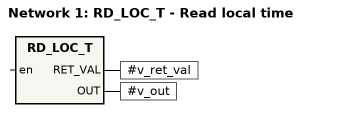
   #v_ret_val := RD_LOC_T(OUT => #v_out);
END_REGION
END_FUNCTION_BLOCK

FUNCTION_BLOCK "FB_Fbd_ex011"   // FB73, FBD
{ S7_Optimized_Access := 'TRUE' }
   VAR_INPUT
      v_req : Bool;
      v_timezone : TimeTransformationRule;
   END_VAR
   VAR_OUTPUT
      v_done : Bool;
      v_busy : Bool;
      v_error : Bool;
      v_status : Word;
   END_VAR
   VAR
      inst : SET_TIMEZONE;
   END_VAR
BEGIN

REGION Network 1: SET_TIMEZONE - Set time zone
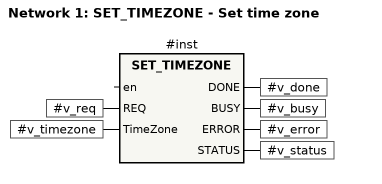
   #inst(REQ := #v_req,   // SET_TIMEZONE
         TimeZone := #v_timezone,
         DONE => #v_done,
         BUSY => #v_busy,
         ERROR => #v_error,
         STATUS => #v_status);
END_REGION
END_FUNCTION_BLOCK

FUNCTION_BLOCK "FB_Fbd_ex012"   // FB74, FBD
{ S7_Optimized_Access := 'TRUE' }
   VAR_OUTPUT
      v_ret_val : Int;
   END_VAR
BEGIN

REGION Network 1: SNC_RTCB - Synchronize slave clocks
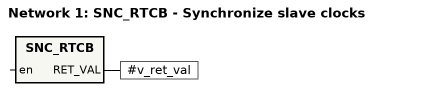
   #v_ret_val := SNC_RTCB();
END_REGION
END_FUNCTION_BLOCK

FUNCTION_BLOCK "FB_Fbd_ex013"   // FB75, FBD
{ S7_Optimized_Access := 'TRUE' }
   VAR_OUTPUT
      v_ret_val : Time;
   END_VAR
BEGIN

REGION Network 1: TIME_TCK - Read time counter
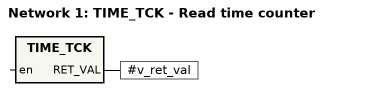
   #v_ret_val := TIME_TCK();
END_REGION
END_FUNCTION_BLOCK

FUNCTION_BLOCK "FB_Fbd_ex014"   // FB76, FBD
{ S7_Optimized_Access := 'TRUE' }
   VAR_INPUT
      v_nr : Rtm;
      v_mode : Byte;
      v_pv : DInt;
   END_VAR
   VAR_OUTPUT
      v_ret_val : Int;
      v_cq : Bool;
      v_cv : DInt;
   END_VAR
BEGIN

REGION Network 1: RTM - Runtime meters
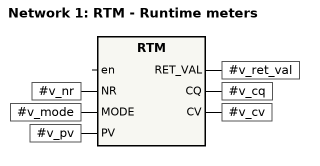
   #v_ret_val := RTM(NR := #v_nr, MODE := #v_mode, PV := #v_pv, CQ => #v_cq, CV => #v_cv);
END_REGION
END_FUNCTION_BLOCK

FUNCTION_BLOCK "FB_Fbd_ex015"   // FB77, FBD
{ S7_Optimized_Access := 'TRUE' }
   VAR_INPUT
      v_in : String;
   END_VAR
   VAR_OUTPUT
      v_out : String;
   END_VAR
BEGIN

REGION Network 1: S_MOVE - Move character string
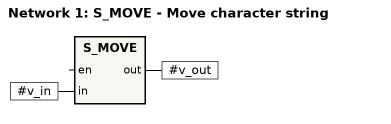
   #v_out := #v_in;
END_REGION
END_FUNCTION_BLOCK

FUNCTION_BLOCK "FB_Fbd_ex025"   // FB78, FBD
{ S7_Optimized_Access := 'TRUE' }
   VAR_INPUT
      v_n : Int;
   END_VAR
   VAR_OUTPUT
      v_ret_val : Word;
   END_VAR
   VAR_IN_OUT
      v_in : Variant;
      v_out : Variant;
   END_VAR
BEGIN

REGION Network 1: ATH - Convert ASCII string to hexadecimal number
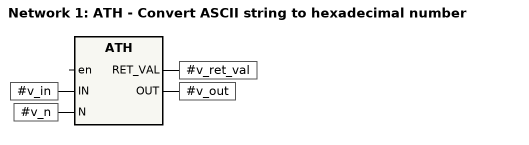
   #v_ret_val := ATH(IN := #v_in, N := #v_n, OUT => #v_out);
END_REGION
END_FUNCTION_BLOCK

FUNCTION_BLOCK "FB_Fbd_ex026"   // FB79, FBD
{ S7_Optimized_Access := 'TRUE' }
   VAR_INPUT
      v_n : UInt;
   END_VAR
   VAR_OUTPUT
      v_ret_val : Word;
   END_VAR
   VAR_IN_OUT
      v_in : Variant;
      v_out : Variant;
   END_VAR
BEGIN

REGION Network 1: HTA - Convert hexadecimal number to ASCII string
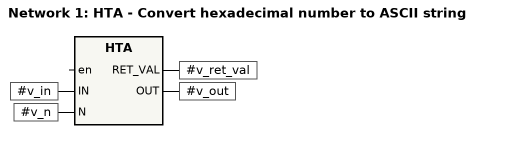
   #v_ret_val := HTA(IN := #v_in, N := #v_n, OUT => #v_out);
END_REGION
END_FUNCTION_BLOCK

FUNCTION_BLOCK "FB_Fbd_ex036"   // FB80, FBD
{ S7_Optimized_Access := 'TRUE' }
   VAR_INPUT
      v_size : DInt;
   END_VAR
   VAR_OUTPUT
      v_out : WString;
   END_VAR
   VAR_IN_OUT
      v_variable : Variant;
   END_VAR
BEGIN

REGION Network 1: GetSymbolName - Read out a tag on the input parameter
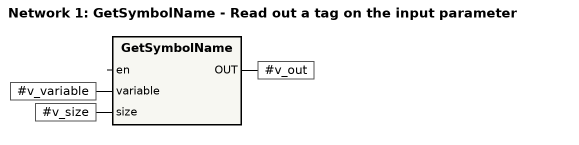
   // no SCL statement known for GetSymbolName: written as a call
   #v_out := GetSymbolName(variable := #v_variable, size := #v_size);
END_REGION
END_FUNCTION_BLOCK

FUNCTION_BLOCK "FB_Fbd_ex038"   // FB81, FBD
{ S7_Optimized_Access := 'TRUE' }
   VAR_INPUT
      v_size : DInt;
   END_VAR
   VAR_OUTPUT
      v_out : WString;
   END_VAR
BEGIN

REGION Network 1: GetInstanceName - Read out name of the read instance
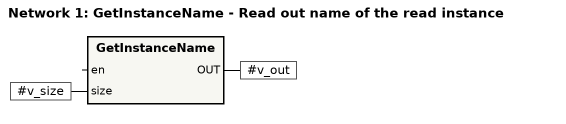
   // no SCL statement known for GetInstanceName: written as a call
   #v_out := GetInstanceName(size := #v_size);
END_REGION
END_FUNCTION_BLOCK

FUNCTION_BLOCK "FB_Fbd_ex039"   // FB82, FBD
{ S7_Optimized_Access := 'TRUE' }
   VAR_INPUT
      v_size : DInt;
   END_VAR
   VAR_OUTPUT
      v_out : WString;
   END_VAR
BEGIN

REGION Network 1: GetInstancePath - Query composite global name of the block instance
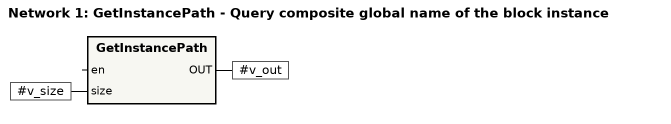
   // no SCL statement known for GetInstancePath: written as a call
   #v_out := GetInstancePath(size := #v_size);
END_REGION
END_FUNCTION_BLOCK

FUNCTION_BLOCK "FB_Fbd_ex040"   // FB83, FBD
{ S7_Optimized_Access := 'TRUE' }
   VAR_INPUT
      v_size : DInt;
   END_VAR
   VAR_OUTPUT
      v_ret_val : WString;
   END_VAR
BEGIN

REGION Network 1: GetBlockName - Read out name of the block
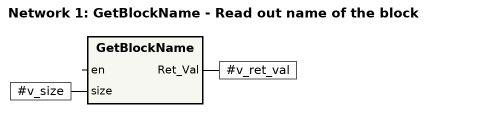
   // no SCL statement known for GetBlockName: written as a call
   #v_ret_val := GetBlockName(size := #v_size);
END_REGION
END_FUNCTION_BLOCK

FUNCTION_BLOCK "FB_Fbd_ex041"   // FB84, FBD
{ S7_Optimized_Access := 'TRUE' }
   VAR_INPUT
      v_part : Pip;
   END_VAR
   VAR_OUTPUT
      v_ret_val : Int;
      v_fladdr : Word;
   END_VAR
BEGIN

REGION Network 1: UPDAT_PI - Update the process image inputs
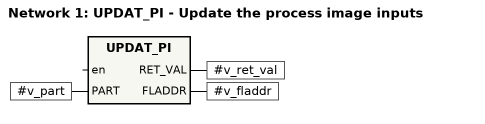
   #v_ret_val := UPDAT_PI(PART := #v_part, FLADDR => #v_fladdr);
END_REGION
END_FUNCTION_BLOCK

FUNCTION_BLOCK "FB_Fbd_ex042"   // FB85, FBD
{ S7_Optimized_Access := 'TRUE' }
   VAR_INPUT
      v_part : Pip;
   END_VAR
   VAR_OUTPUT
      v_ret_val : Int;
      v_fladdr : Word;
   END_VAR
BEGIN

REGION Network 1: UPDAT_PO - Update the process image outputs
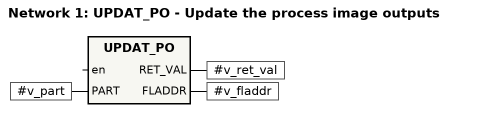
   #v_ret_val := UPDAT_PO(PART := #v_part, FLADDR => #v_fladdr);
END_REGION
END_FUNCTION_BLOCK

FUNCTION_BLOCK "FB_Fbd_ex043"   // FB86, FBD
{ S7_Optimized_Access := 'TRUE' }
   VAR_INPUT
      v_part : Pip;
   END_VAR
   VAR_OUTPUT
      v_ret_val : Int;
      v_fladdr : Word;
   END_VAR
BEGIN

REGION Network 1: SYNC_PI - Synchronize the process image inputs
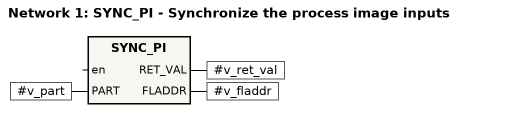
   #v_ret_val := SYNC_PI(PART := #v_part, FLADDR => #v_fladdr);
END_REGION
END_FUNCTION_BLOCK

FUNCTION_BLOCK "FB_Fbd_ex044"   // FB87, FBD
{ S7_Optimized_Access := 'TRUE' }
   VAR_INPUT
      v_part : Pip;
   END_VAR
   VAR_OUTPUT
      v_ret_val : Int;
      v_fladdr : Word;
   END_VAR
BEGIN

REGION Network 1: SYNC_PO - Synchronize the process image outputs
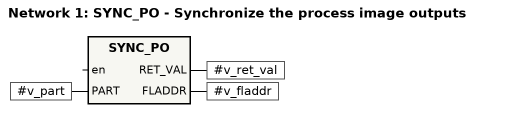
   #v_ret_val := SYNC_PO(PART := #v_part, FLADDR => #v_fladdr);
END_REGION
END_FUNCTION_BLOCK

FUNCTION_BLOCK "FB_Fbd_ex045"   // FB88, FBD
{ S7_Optimized_Access := 'TRUE' }
   VAR_INPUT
      v_req : Bool;
      v_id : Hw_Io;
      v_index : DInt;
      v_mlen : UInt;
   END_VAR
   VAR_OUTPUT
      v_valid : Bool;
      v_busy : Bool;
      v_error : Bool;
      v_status : DWord;
      v_len : UInt;
   END_VAR
   VAR_IN_OUT
      v_record : Array[0..99] of Byte;
   END_VAR
   VAR
      inst : RDREC;
   END_VAR
BEGIN

REGION Network 1: RDREC - Read data record
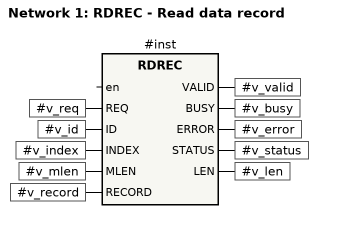
   #inst(REQ := #v_req,   // RDREC
         ID := #v_id,
         INDEX := #v_index,
         MLEN := #v_mlen,
         RECORD := #v_record,
         VALID => #v_valid,
         BUSY => #v_busy,
         ERROR => #v_error,
         STATUS => #v_status,
         LEN => #v_len);
END_REGION
END_FUNCTION_BLOCK

FUNCTION_BLOCK "FB_Fbd_ex046"   // FB89, FBD
{ S7_Optimized_Access := 'TRUE' }
   VAR_INPUT
      v_req : Bool;
      v_id : Hw_Io;
      v_index : DInt;
      v_len : UInt;
   END_VAR
   VAR_OUTPUT
      v_done : Bool;
      v_busy : Bool;
      v_error : Bool;
      v_status : DWord;
   END_VAR
   VAR_IN_OUT
      v_record : Array[0..99] of Byte;
   END_VAR
   VAR
      inst : WRREC;
   END_VAR
BEGIN

REGION Network 1: WRREC - Write data record
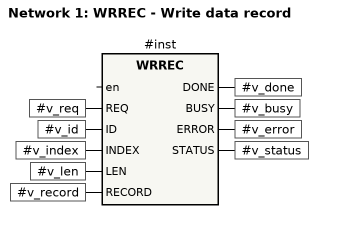
   #inst(REQ := #v_req,   // WRREC
         ID := #v_id,
         INDEX := #v_index,
         LEN := #v_len,
         RECORD := #v_record,
         DONE => #v_done,
         BUSY => #v_busy,
         ERROR => #v_error,
         STATUS => #v_status);
END_REGION
END_FUNCTION_BLOCK

FUNCTION_BLOCK "FB_Fbd_ex047"   // FB90, FBD
{ S7_Optimized_Access := 'TRUE' }
   VAR_INPUT
      v_id : Hw_SubModule;
   END_VAR
   VAR_OUTPUT
      v_status : DWord;
      v_len : Int;
   END_VAR
   VAR_IN_OUT
      v_inputs : Array[0..99] of Byte;
   END_VAR
   VAR
      inst : GETIO;
   END_VAR
BEGIN

REGION Network 1: GETIO - Read all inputs of a submodule
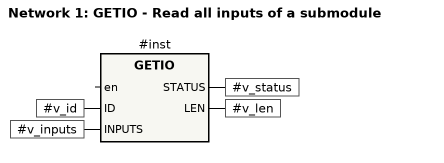
   #inst(ID := #v_id, INPUTS := #v_inputs, STATUS => #v_status, LEN => #v_len);   // GETIO
END_REGION
END_FUNCTION_BLOCK

FUNCTION_BLOCK "FB_Fbd_ex048"   // FB91, FBD
{ S7_Optimized_Access := 'TRUE' }
   VAR_INPUT
      v_id : Hw_SubModule;
   END_VAR
   VAR_OUTPUT
      v_status : DWord;
   END_VAR
   VAR_IN_OUT
      v_outputs : Array[0..99] of Byte;
   END_VAR
   VAR
      inst : SETIO;
   END_VAR
BEGIN

REGION Network 1: SETIO - Write all outputs of a submodule
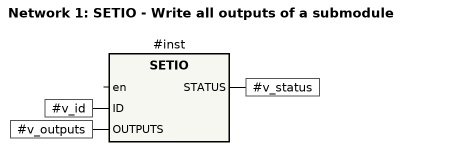
   #inst(ID := #v_id, OUTPUTS := #v_outputs, STATUS => #v_status);   // SETIO
END_REGION
END_FUNCTION_BLOCK

FUNCTION_BLOCK "FB_Fbd_ex049"   // FB92, FBD
{ S7_Optimized_Access := 'TRUE' }
   VAR_INPUT
      v_id : Hw_SubModule;
      v_offset : Int;
      v_len : Int;
   END_VAR
   VAR_OUTPUT
      v_status : DWord;
      v_error : Bool;
   END_VAR
   VAR_IN_OUT
      v_inputs : Array[0..99] of Byte;
   END_VAR
   VAR
      inst : GETIO_PART;
   END_VAR
BEGIN

REGION Network 1: GETIO_PART - Read inputs of a submodule
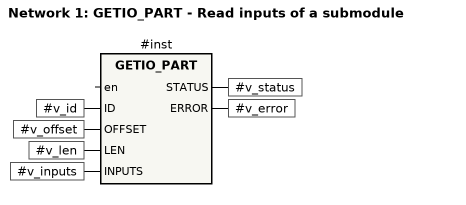
   #inst(ID := #v_id,   // GETIO_PART
         OFFSET := #v_offset,
         LEN := #v_len,
         INPUTS := #v_inputs,
         STATUS => #v_status,
         ERROR => #v_error);
END_REGION
END_FUNCTION_BLOCK

FUNCTION_BLOCK "FB_Fbd_ex050"   // FB93, FBD
{ S7_Optimized_Access := 'TRUE' }
   VAR_INPUT
      v_id : Hw_SubModule;
      v_offset : Int;
      v_len : Int;
   END_VAR
   VAR_OUTPUT
      v_status : DWord;
      v_error : Bool;
   END_VAR
   VAR_IN_OUT
      v_outputs : Array[0..99] of Byte;
   END_VAR
   VAR
      inst : SETIO_PART;
   END_VAR
BEGIN

REGION Network 1: SETIO_PART - Write outputs of a submodule
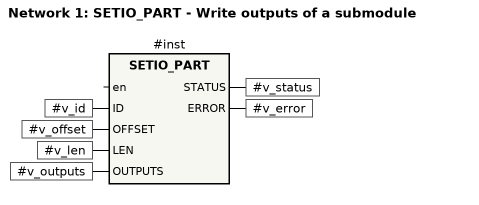
   #inst(ID := #v_id,   // SETIO_PART
         OFFSET := #v_offset,
         LEN := #v_len,
         OUTPUTS := #v_outputs,
         STATUS => #v_status,
         ERROR => #v_error);
END_REGION
END_FUNCTION_BLOCK

FUNCTION_BLOCK "FB_Fbd_ex056"   // FB94, FBD
{ S7_Optimized_Access := 'TRUE' }
   VAR_INPUT
      v_req : Bool;
      v_mode : USInt;
      v_laddr : Hw_Device;
   END_VAR
   VAR_OUTPUT
      v_ret_val : Int;
      v_busy : Bool;
   END_VAR
BEGIN

REGION Network 1: D_ACT_DP - Activate/deactivate DP slaves
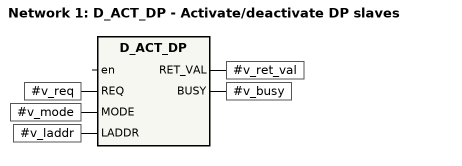
   #v_ret_val := D_ACT_DP(REQ := #v_req, MODE := #v_mode, LADDR := #v_laddr, BUSY => #v_busy);
END_REGION
END_FUNCTION_BLOCK

FUNCTION_BLOCK "FB_Fbd_ex057"   // FB95, FBD
{ S7_Optimized_Access := 'TRUE' }
   VAR_INPUT
      v_req : Bool;
      v_mode : UInt;
      v_laddr : Hw_Interface;
      v_ctrlrec : Array[0..99] of Byte;
   END_VAR
   VAR_OUTPUT
      v_done : Bool;
      v_busy : Bool;
      v_error : Bool;
      v_status : DWord;
      v_err_info : Word;
   END_VAR
   VAR
      inst : ReconfigIOSystem;
   END_VAR
BEGIN

REGION Network 1: ReconfigIOSystem - Reconfigure IO system
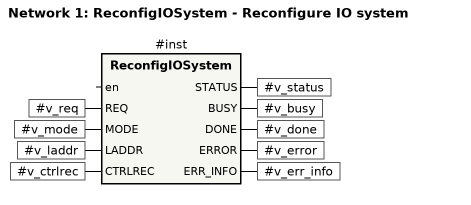
   #inst(REQ := #v_req,   // ReconfigIOSystem
         MODE := #v_mode,
         LADDR := #v_laddr,
         CTRLREC := #v_ctrlrec,
         STATUS => #v_status,
         BUSY => #v_busy,
         DONE => #v_done,
         ERROR => #v_error,
         ERR_INFO => #v_err_info);
END_REGION
END_FUNCTION_BLOCK

FUNCTION_BLOCK "FB_Fbd_ex060"   // FB96, FBD
{ S7_Optimized_Access := 'TRUE' }
   VAR_INPUT
      v_laddr : Hw_Io;
   END_VAR
   VAR_OUTPUT
      v_ret_val : Int;
   END_VAR
   VAR_IN_OUT
      v_record : Variant;
   END_VAR
BEGIN

REGION Network 1: DPRD_DAT - Read consistent data of a DP standard slave
